// This function has been automatically generated from the project information.
{attribute 'signature_flag' := '1073741824'}
{attribute 'TcGenerated'}
{attribute 'no-analysis'}
FUNCTION F_GetTitle : WSTRING
VAR_INPUT
	
END_VAR

F_GetTitle := "TcOtlp";

END_FUNCTION

(* stored: Version 1.1.0.1
   POU F_GetTitle: Id {92df87f7-baa6-46e4-ac51-b3d27789699d}, SpecialFunc None *)
